FUNCTION_BLOCK AOption_AD_DEMUX_4 (* AOption Bitmasken-Demultiplexor (generic FB): aktiviert per Bitmaske K beliebig viele von 4 Options-Ausgaengen (INIT_REQ), Multi-Select. *)
  (* Standard: 61499-2; Description: Copyright (c) 2026 Meisterschulen am Ostbahnhof This program and the accompanying materials are made available under the terms of the Eclipse Public License 2.0 which is available at https://www.eclipse.org/legal/epl-2.0/ SPDX-License-Identifier: EPL-2.0 *)
  (* Version 1.0, 2026-10-13, Franz Höpfinger, Meisterschulen am Ostbahnhof *)
  PACKAGE Option::selection;
  {SET_ATTRIBUTE(eclipse4diac::core::GenericClassName, 'GEN_AOption_AD_DEMUX')}
  (* Documentation:
  Demultiplexer (natives Generic-FB, kein ECC/Algorithmus in diesem Typ) fuer N=4 Options-Ausgaenge vom Typ Option::AOption, ausgewaehlt ueber den bidirektionalen Bitmasken-Adapter K (adapter::types::bidirectional::AD2, DWORD).
   Bitzuordnung (Multi-Select, im Gegensatz zum Single-Select von AOption_AUI_DEMUX_4):
    - Bit 0 (Wert 1) – OUT1
   - Bit 1 (Wert 2) – OUT2
   - Bit 2 (Wert 4) – OUT3
   - Bit 3 (Wert 8) – OUT4
    Beispiel: K = 3 (Bit 0 + Bit 1 gesetzt) – OUT1 UND OUT2 an, alle anderen aus. Es koennen beliebig viele bzw. alle Ausgaenge gleichzeitig aktiv sein.
   Umschaltverhalten: nur Bits, die sich gegenueber dem vorherigen K-Wert aendern, loesen an dem zugehoerigen Ausgang ein INIT_REQ aus (0→1: QI=TRUE aktivieren, 1→0: QI=FALSE deaktivieren). Unveraenderte Bits werden nicht erneut getriggert - jeder Ausgang wird also pro eintreffendem K-Wert maximal 1x getriggert.
   Busy-Gating ueber den bidirektionalen K-Adapter: Waehrend noch auf INIT_CNF von mindestens einem durch den letzten K-Wechsel betroffenen Ausgang gewartet wird, wird jeder weitere ueber K (Richtung Plug -> Socket, EO1/DO1) eintreffende Bitmasken-Wunsch ignoriert - er wird weder gepuffert noch nachgeholt. Erst wenn alle durch den letzten Wechsel ausgeloesten INIT_CNF eingetroffen sind, meldet der DEMUX dies rueckwaerts ueber K (Richtung Socket -> Plug, EI1/DI1) mit der uebernommenen Bitmaske zurueck (nicht mit dem Zustand der Ausgaenge: auch Bits ausserhalb der vorhandenen Ausgaenge werden unveraendert quittiert); erst danach werden wieder neue K-Wuensche angenommen. Damit sind sowohl langsame Umschaltvorgaenge als auch mehrfache, einander widersprechende K-Werte in kurzer Folge sauber abgedeckt.
  *)
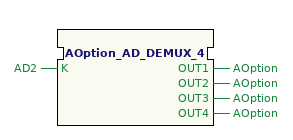
  SOCKETS
    K : adapter::types::bidirectional::AD2; (* Bitmaske (Bit0=OUT1, Bit1=OUT2, ...), bidirektional: EO1/DO1 = neuer Bitmasken-Wunsch rein, EI1/DI1 = Quittung mit der uebernommenen Bitmaske zurueck *)
  END_SOCKETS
  PLUGS
    OUT1 : Option::AOption; (* Option 1 (aktiv wenn Bit 0 von K gesetzt ist, Wert 1) *)
    OUT2 : Option::AOption; (* Option 2 (aktiv wenn Bit 1 von K gesetzt ist, Wert 2) *)
    OUT3 : Option::AOption; (* Option 3 (aktiv wenn Bit 2 von K gesetzt ist, Wert 4) *)
    OUT4 : Option::AOption; (* Option 4 (aktiv wenn Bit 3 von K gesetzt ist, Wert 8) *)
  END_PLUGS
END_FUNCTION_BLOCK
